(* IEC 61131-3 sources: plc-ci-toolkit/ci/tests/samples/sa_probe_src/src/POUs/F_SaTemp, 1 file *)

(* ---- F_SaTemp.decl.st ---- *)
// Назначение: зонд статанализа (намеренно плохой код)
{attribute 'analysis' := '-167'}
FUNCTION F_SaTemp : BOOL
VAR_INPUT
    xIn : BOOL;
END_VAR
VAR
    fbDelay : FB_Example;           // SA0167: временный экземпляр ФБ в функции
END_VAR
